PROGRAM prg_RecipeManager
VAR
	fbRecipe: RecipeManCommands;
	LastError: DWORD;
	LastInfo: InfoValues;

	bCheckError: BOOL;
	bResetError: BOOL;
	bInit: BOOL;
END_VAR


IF bCheckError THEN;
	//bCheckError:=FALSE;
	LastError:=fbRecipe.GetLastError();
	LastInfo:=fbRecipe.GetLastInfo();
END_IF

IF bResetError THEN;
	bResetError:=FALSE;
	LastError:=fbRecipe.ResetLastError();
	LastError:=fbRecipe.ReloadRecipes(RecipeDefinitionName:='');
	
END_IF

IF bInit THEN;
	bInit:=FALSE;
	LastError:=fbRecipe.ResetLastInfo();
END_IF

END_PROGRAM

(* stored: Version 1.1.0.1, ProductVersion 3.1.4024.12
   POU prg_RecipeManager: Id {85473640-566c-4030-8ff1-15160df57023}, SpecialFunc None *)
